FUNCTION_BLOCK GcfFunctionCallTest (* Test: F_Double ueber GCF und direkt aufrufen *)
  (* Standard: 61499-1; Description: Copyright (c) 2026 Meisterschulen am Ostbahnhof This program and the accompanying materials are made available under the terms of the Eclipse Public License 2.0 which is available at https://www.eclipse.org/legal/epl-2.0/ SPDX-License-Identifier: EPL-2.0 *)
  (* Version 1.0, 2026-10-16, Franz Höpfinger, Meisterschulen am Ostbahnhof, Uebung: Function aus GCF aufrufen *)
  PACKAGE Meins::GcfFunctionCall;
  IMPORT Meins::GcfFunctionCall::const::FuncConst::DOUBLE_VALUE;
  IMPORT Meins::GcfFunctionCall::const::FuncConst::BASE_VALUE;
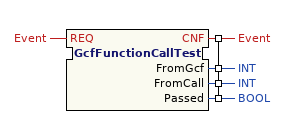
  EVENT_INPUT
    REQ;
  END_EVENT
  EVENT_OUTPUT
    CNF WITH FromGcf, FromCall, Passed;
  END_EVENT
  VAR_OUTPUT
    FromGcf : INT; (* DOUBLE_VALUE aus GCF *)
    FromCall : INT; (* F_Double direkt im ST *)
    Passed : BOOL; (* TRUE wenn beide 14 *)
  END_VAR
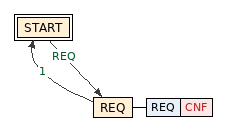
  EC_STATES
    START; (* Initial State *)
    REQ : REQ -> CNF; (* Normal execution *)
  END_STATES
  EC_TRANSITIONS
    START TO REQ := REQ;
    REQ TO START := 1;
  END_TRANSITIONS
  ALGORITHM REQ IN ST: (* Normal execution *)
FromGcf := DOUBLE_VALUE;
FromCall := Meins::GcfFunctionCall::F_Double(BASE_VALUE);
Passed := (FromGcf = 14) AND (FromCall = 14);
  END_ALGORITHM
END_FUNCTION_BLOCK
